// FB_TP: 脉冲定时器
// 描述: 当IN上升沿时, Q输出固定时长PT的脉冲

FUNCTION_BLOCK FB_TP
VAR_INPUT
    IN  : BOOL;
    PT  : DINT;   // 脉冲宽度(扫描周期)
END_VAR
VAR_OUTPUT
    Q   : BOOL;
    ET  : DINT;   // 已用时间(扫描周期)
END_VAR
VAR
    Counter   : DINT := 0;
    Running   : BOOL := FALSE;
END_VAR

BEGIN
    // 检测IN上升沿
    IF #IN AND NOT #Running THEN
        #Running := TRUE;
        #Counter := 0;
        #Q := TRUE;
    END_IF;

    // 脉冲计时
    IF #Running THEN
        #Counter := #Counter + 1;
        #ET := #Counter;

        IF #Counter >= #PT THEN
            #Q := FALSE;
            #Running := FALSE;
        END_IF;
    ELSIF NOT #IN THEN
        #Q := FALSE;
        #ET := 0;
        #Counter := 0;
    END_IF;

END_FUNCTION_BLOCK
